FUNCTION CheckDivReal_1 : REAL
VAR_INPUT
	divisor: REAL;
END_VAR
VAR_EXTERNAL
	fbCheckDivRealInfo: FB_CheckDivRealInfo;
END_VAR

(*This function checks if a division by zero is performed*)

fbCheckDivRealInfo(
	rDivisor			:= divisor,
	sLogMessage	=> ,
	rReturnDivReal 	=> CheckDivReal);

END_FUNCTION

(* stored: Version 1.1.0.1, ProductVersion 3.1.4024.15
   POU CheckDivReal_1: Id {e50bf1c7-8480-4e31-aba5-bdfe3a40881e}, SpecialFunc CheckDivReal32 *)
